SYSTEM SINF_0
  (* Version 1.0, 2023-02-20, eliseu *)
  APPLICATION SINF_0App
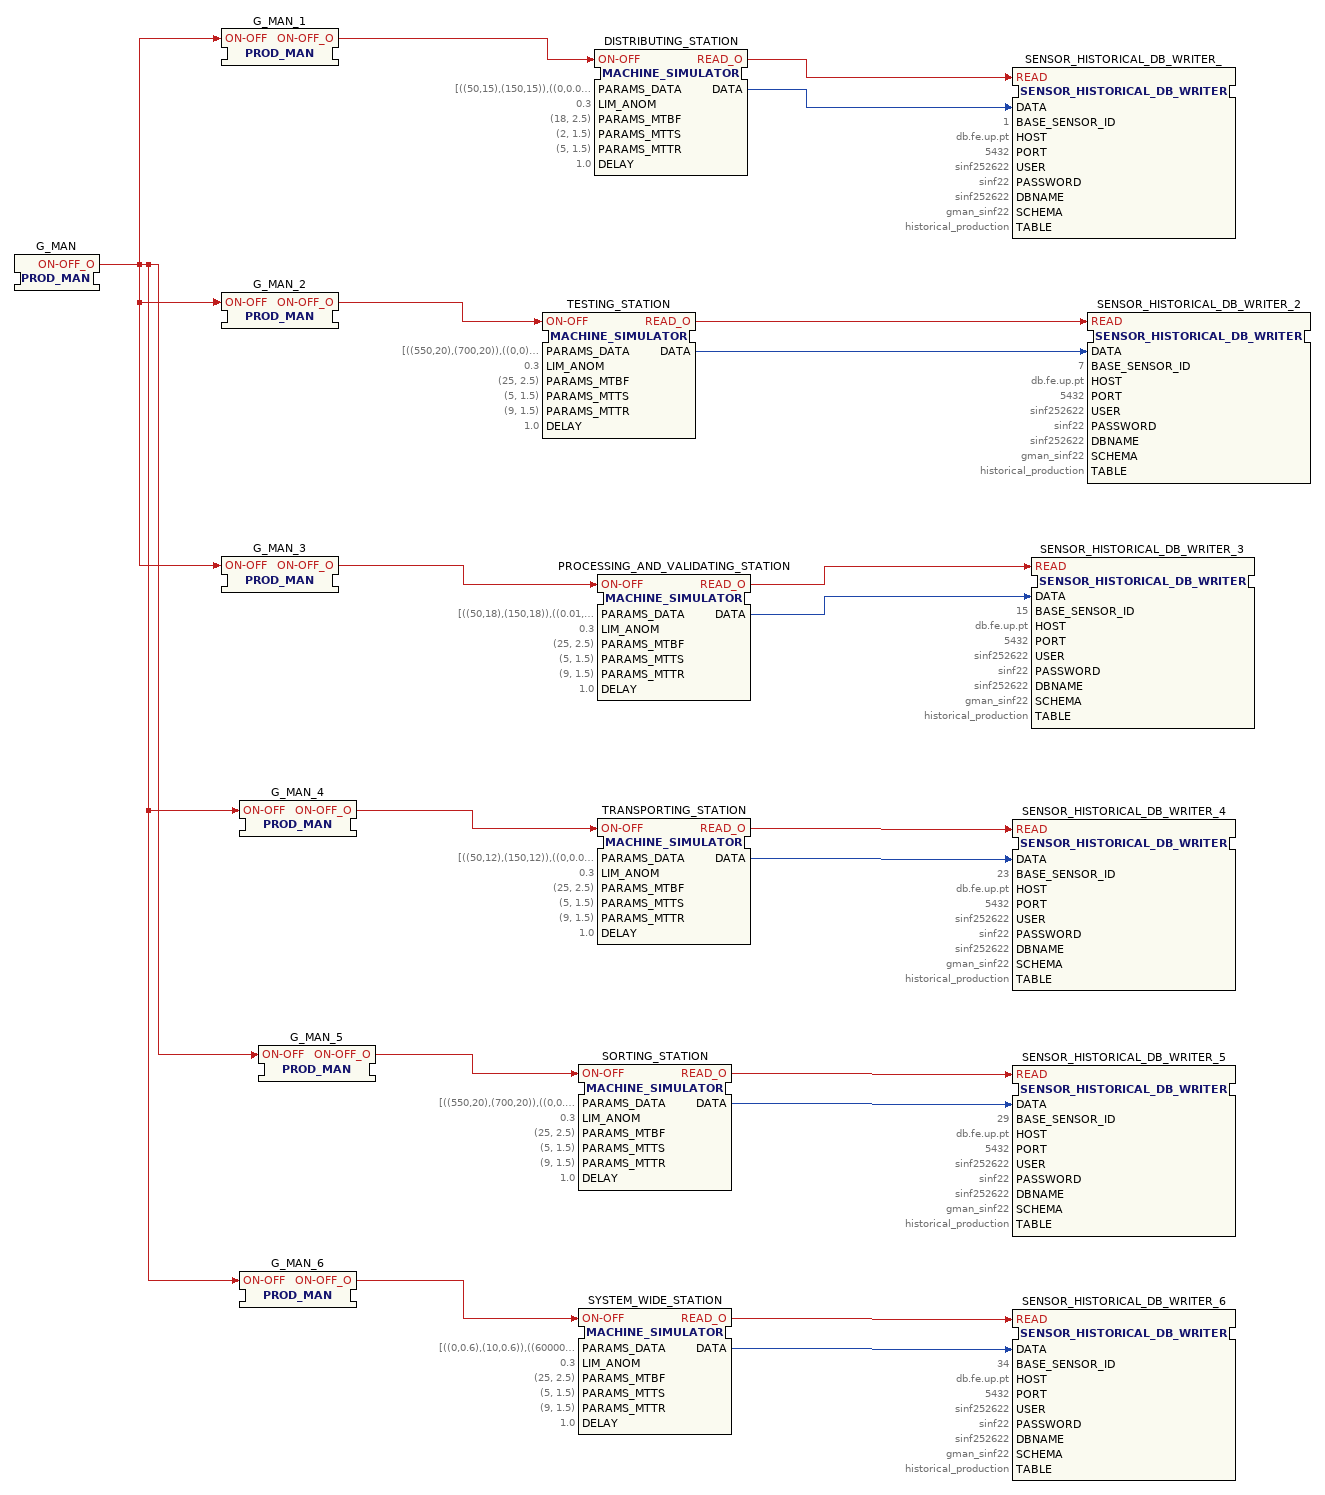
    FBS
      G_MAN_1 : PROD_MAN;
      DISTRIBUTING_STATION : MACHINE_SIMULATOR(PARAMS_DATA := [((50,15),(150,15)),((0,0.05),(3,0.05)),((600000,30000),(800000,30000)),((0.01,0.008),(0.05,0.008)),((2,0.4),(5,0.4)),((293,2.5),(303,2.5))], LIM_ANOM := 0.3, PARAMS_MTBF := (18, 2.5), PARAMS_MTTS := (2, 1.5), PARAMS_MTTR := (5, 1.5), DELAY := 1.0);
      TESTING_STATION : MACHINE_SIMULATOR(PARAMS_DATA := [((550,20),(700,20)),((0,0),(1,0)),((0.2,0.12),(0.8,0.12)),((0,0.05),(3,0.05)),((300,120),(1000,120)),((40,5),(60,5)),((293,2.5),(303,2.5)),((0,0.3),(2,0.3))], LIM_ANOM := 0.3, PARAMS_MTBF := (25, 2.5), PARAMS_MTTS := (5, 1.5), PARAMS_MTTR := (9, 1.5), DELAY := 1.0);
      PROCESSING_AND_VALIDATING_STATION : MACHINE_SIMULATOR(PARAMS_DATA := [((50,18),(150,18)),((0.01,0.012),(0.1,0.012)),((0,0),(1,0)),((0,0.05),(3,0.05)),((2,0.4),(5,0.4)),((333,6),(353,6)),((0.01,0.007),(0.05,0.007)),((500,100),(1000,100))], LIM_ANOM := 0.3, PARAMS_MTBF := (25, 2.5), PARAMS_MTTS := (5, 1.5), PARAMS_MTTR := (9, 1.5), DELAY := 1.0);
      TRANSPORTING_STATION : MACHINE_SIMULATOR(PARAMS_DATA := [((50,12),(150,12)),((0,0.05),(3,0.05)),((2,0.4),(5,0.4)),((333,5),(333,5)),((600000,25000),(800000,25000)),((0.01,0.006),(0.05,0.006))], LIM_ANOM := 0.3, PARAMS_MTBF := (25, 2.5), PARAMS_MTTS := (5, 1.5), PARAMS_MTTR := (9, 1.5), DELAY := 1.0);
      SORTING_STATION : MACHINE_SIMULATOR(PARAMS_DATA := [((550,20),(700,20)),((0,0.05),(3,0.05)),((300,150),(1000,150)),((2,0.35),(5,0.35)),((293,2.5),(303,2.5))], LIM_ANOM := 0.3, PARAMS_MTBF := (25, 2.5), PARAMS_MTTS := (5, 1.5), PARAMS_MTTR := (9, 1.5), DELAY := 1.0);
      SYSTEM_WIDE_STATION : MACHINE_SIMULATOR(PARAMS_DATA := [((0,0.6),(10,0.6)),((600000,30000),(800000,30000)),((40,5),(60,5)),((293,2.5),(303,2.5))], LIM_ANOM := 0.3, PARAMS_MTBF := (25, 2.5), PARAMS_MTTS := (5, 1.5), PARAMS_MTTR := (9, 1.5), DELAY := 1.0);
      G_MAN_2 : PROD_MAN;
      G_MAN_3 : PROD_MAN;
      G_MAN_4 : PROD_MAN;
      G_MAN_5 : PROD_MAN;
      G_MAN_6 : PROD_MAN;
      G_MAN : PROD_MAN;
      SENSOR_HISTORICAL_DB_WRITER_ : SENSOR_HISTORICAL_DB_WRITER(BASE_SENSOR_ID := 1, HOST := db.fe.up.pt, PORT := 5432, USER := sinf252622, PASSWORD := sinf22, DBNAME := sinf252622, SCHEMA := gman_sinf22, TABLE := historical_production);
      SENSOR_HISTORICAL_DB_WRITER_2 : SENSOR_HISTORICAL_DB_WRITER(BASE_SENSOR_ID := 7, HOST := db.fe.up.pt, PORT := 5432, USER := sinf252622, PASSWORD := sinf22, DBNAME := sinf252622, SCHEMA := gman_sinf22, TABLE := historical_production);
      SENSOR_HISTORICAL_DB_WRITER_3 : SENSOR_HISTORICAL_DB_WRITER(BASE_SENSOR_ID := 15, HOST := db.fe.up.pt, PORT := 5432, USER := sinf252622, PASSWORD := sinf22, DBNAME := sinf252622, SCHEMA := gman_sinf22, TABLE := historical_production);
      SENSOR_HISTORICAL_DB_WRITER_4 : SENSOR_HISTORICAL_DB_WRITER(BASE_SENSOR_ID := 23, HOST := db.fe.up.pt, PORT := 5432, USER := sinf252622, PASSWORD := sinf22, DBNAME := sinf252622, SCHEMA := gman_sinf22, TABLE := historical_production);
      SENSOR_HISTORICAL_DB_WRITER_5 : SENSOR_HISTORICAL_DB_WRITER(BASE_SENSOR_ID := 29, HOST := db.fe.up.pt, PORT := 5432, USER := sinf252622, PASSWORD := sinf22, DBNAME := sinf252622, SCHEMA := gman_sinf22, TABLE := historical_production);
      SENSOR_HISTORICAL_DB_WRITER_6 : SENSOR_HISTORICAL_DB_WRITER(BASE_SENSOR_ID := 34, HOST := db.fe.up.pt, PORT := 5432, USER := sinf252622, PASSWORD := sinf22, DBNAME := sinf252622, SCHEMA := gman_sinf22, TABLE := historical_production);
    END_FBS
    EVENT_CONNECTIONS
      G_MAN_1.ON-OFF_O TO DISTRIBUTING_STATION.ON-OFF;
      G_MAN_2.ON-OFF_O TO TESTING_STATION.ON-OFF;
      G_MAN_3.ON-OFF_O TO PROCESSING_AND_VALIDATING_STATION.ON-OFF;
      G_MAN_4.ON-OFF_O TO TRANSPORTING_STATION.ON-OFF;
      G_MAN_5.ON-OFF_O TO SORTING_STATION.ON-OFF;
      G_MAN_6.ON-OFF_O TO SYSTEM_WIDE_STATION.ON-OFF;
      G_MAN.ON-OFF_O TO G_MAN_1.ON-OFF;
      G_MAN.ON-OFF_O TO G_MAN_2.ON-OFF;
      G_MAN.ON-OFF_O TO G_MAN_3.ON-OFF;
      G_MAN.ON-OFF_O TO G_MAN_4.ON-OFF;
      G_MAN.ON-OFF_O TO G_MAN_5.ON-OFF;
      G_MAN.ON-OFF_O TO G_MAN_6.ON-OFF;
      DISTRIBUTING_STATION.READ_O TO SENSOR_HISTORICAL_DB_WRITER_.READ;
      TESTING_STATION.READ_O TO SENSOR_HISTORICAL_DB_WRITER_2.READ;
      SORTING_STATION.READ_O TO SENSOR_HISTORICAL_DB_WRITER_5.READ;
      TRANSPORTING_STATION.READ_O TO SENSOR_HISTORICAL_DB_WRITER_4.READ;
      PROCESSING_AND_VALIDATING_STATION.READ_O TO SENSOR_HISTORICAL_DB_WRITER_3.READ;
      SYSTEM_WIDE_STATION.READ_O TO SENSOR_HISTORICAL_DB_WRITER_6.READ;
    END_CONNECTIONS
    DATA_CONNECTIONS
      DISTRIBUTING_STATION.DATA TO SENSOR_HISTORICAL_DB_WRITER_.DATA;
      TESTING_STATION.DATA TO SENSOR_HISTORICAL_DB_WRITER_2.DATA;
      SORTING_STATION.DATA TO SENSOR_HISTORICAL_DB_WRITER_5.DATA;
      PROCESSING_AND_VALIDATING_STATION.DATA TO SENSOR_HISTORICAL_DB_WRITER_3.DATA;
      SYSTEM_WIDE_STATION.DATA TO SENSOR_HISTORICAL_DB_WRITER_6.DATA;
      TRANSPORTING_STATION.DATA TO SENSOR_HISTORICAL_DB_WRITER_4.DATA;
    END_CONNECTIONS
  END_APPLICATION
  DEVICE FORTE_PC : FORTE_PC(MGR_ID := "localhost:61499")
    {SET_ATTRIBUTE(Profile, HOLOBLOC)} (* device profile *)
    RESOURCE DIN1 : EMB_RES
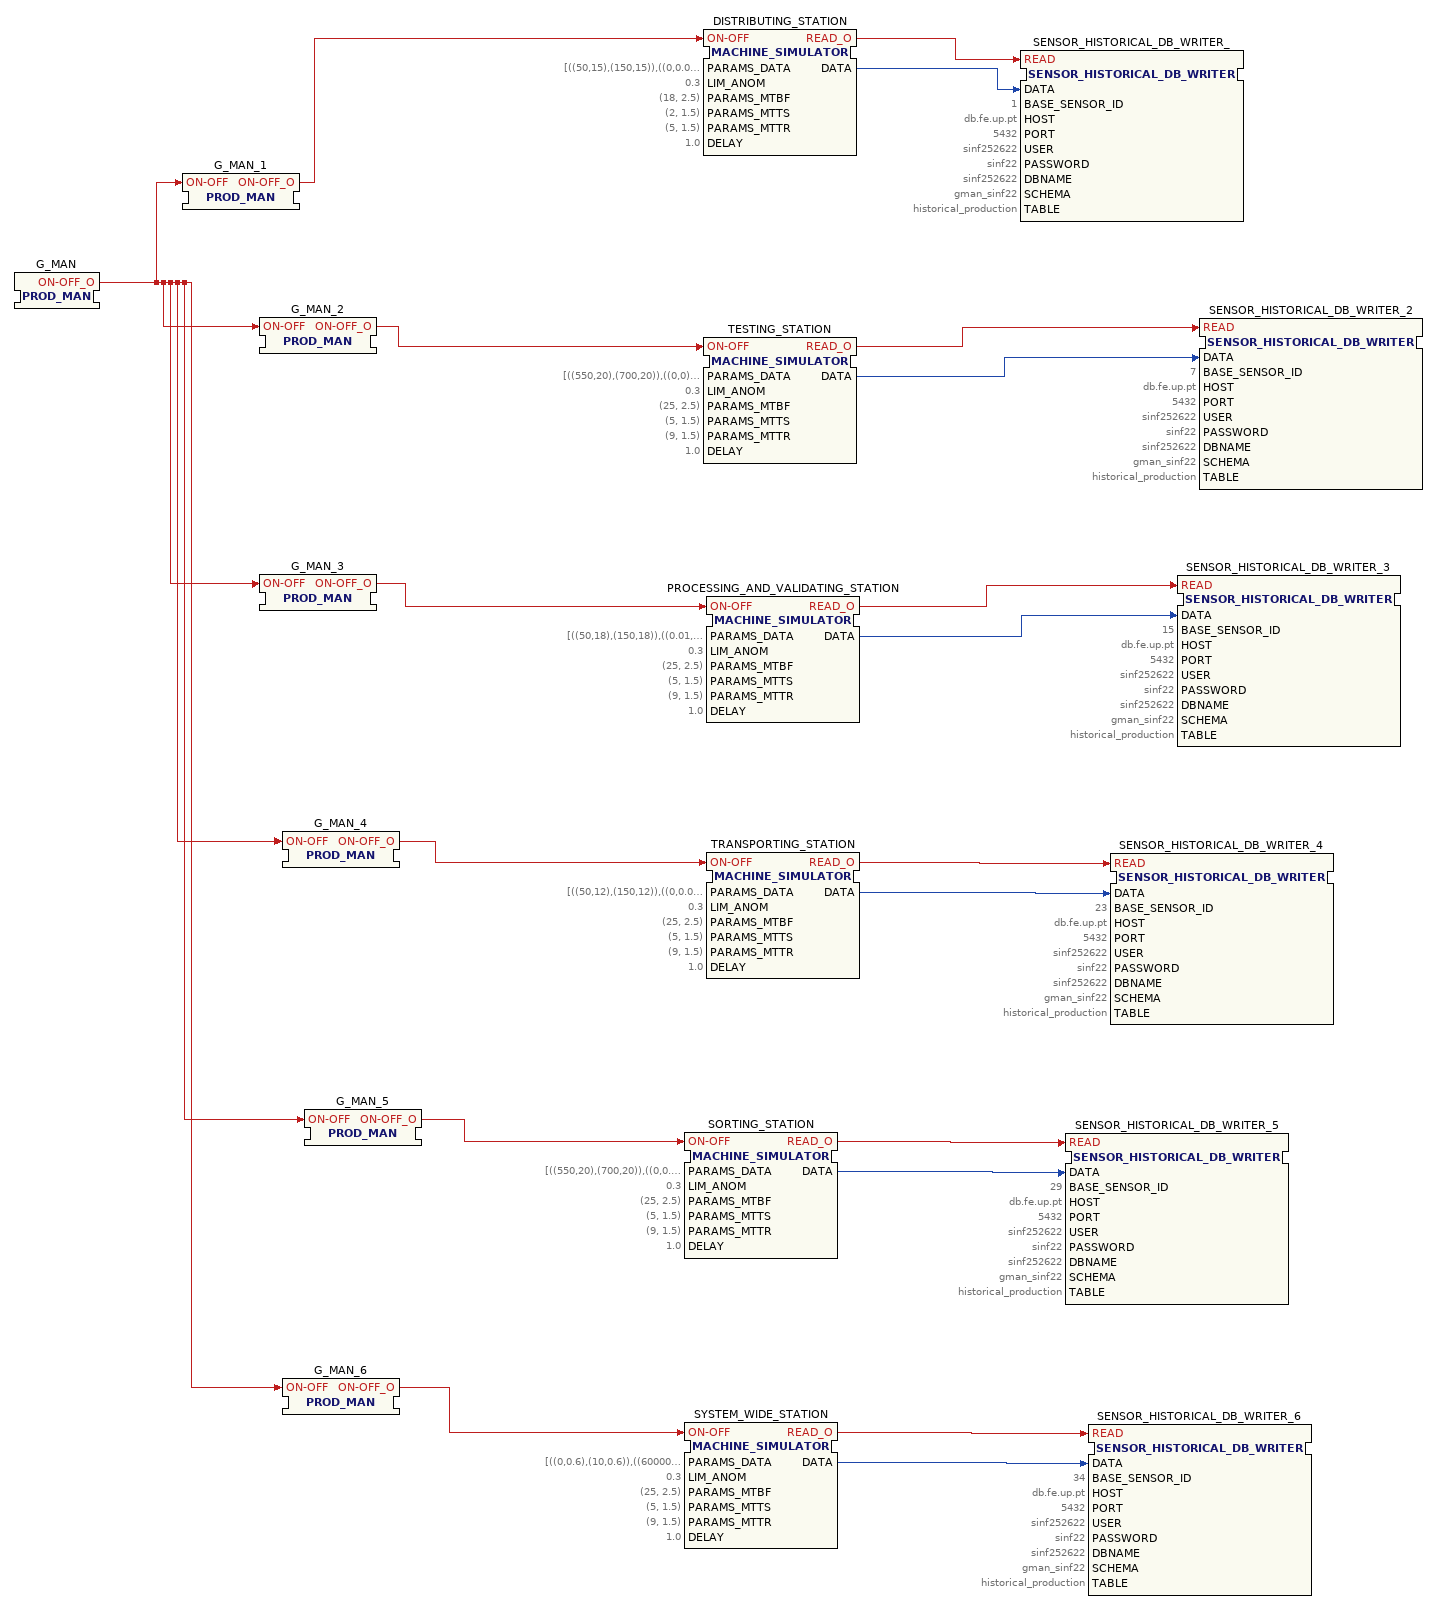
      FBS
        G_MAN_1 : PROD_MAN;
        DISTRIBUTING_STATION : MACHINE_SIMULATOR(PARAMS_DATA := [((50,15),(150,15)),((0,0.05),(3,0.05)),((600000,30000),(800000,30000)),((0.01,0.008),(0.05,0.008)),((2,0.4),(5,0.4)),((293,2.5),(303,2.5))], LIM_ANOM := 0.3, PARAMS_MTBF := (18, 2.5), PARAMS_MTTS := (2, 1.5), PARAMS_MTTR := (5, 1.5), DELAY := 1.0);
        TESTING_STATION : MACHINE_SIMULATOR(PARAMS_DATA := [((550,20),(700,20)),((0,0),(1,0)),((0.2,0.12),(0.8,0.12)),((0,0.05),(3,0.05)),((300,120),(1000,120)),((40,5),(60,5)),((293,2.5),(303,2.5)),((0,0.3),(2,0.3))], LIM_ANOM := 0.3, PARAMS_MTBF := (25, 2.5), PARAMS_MTTS := (5, 1.5), PARAMS_MTTR := (9, 1.5), DELAY := 1.0);
        PROCESSING_AND_VALIDATING_STATION : MACHINE_SIMULATOR(PARAMS_DATA := [((50,18),(150,18)),((0.01,0.012),(0.1,0.012)),((0,0),(1,0)),((0,0.05),(3,0.05)),((2,0.4),(5,0.4)),((333,6),(353,6)),((0.01,0.007),(0.05,0.007)),((500,100),(1000,100))], LIM_ANOM := 0.3, PARAMS_MTBF := (25, 2.5), PARAMS_MTTS := (5, 1.5), PARAMS_MTTR := (9, 1.5), DELAY := 1.0);
        TRANSPORTING_STATION : MACHINE_SIMULATOR(PARAMS_DATA := [((50,12),(150,12)),((0,0.05),(3,0.05)),((2,0.4),(5,0.4)),((333,5),(333,5)),((600000,25000),(800000,25000)),((0.01,0.006),(0.05,0.006))], LIM_ANOM := 0.3, PARAMS_MTBF := (25, 2.5), PARAMS_MTTS := (5, 1.5), PARAMS_MTTR := (9, 1.5), DELAY := 1.0);
        SORTING_STATION : MACHINE_SIMULATOR(PARAMS_DATA := [((550,20),(700,20)),((0,0.05),(3,0.05)),((300,150),(1000,150)),((2,0.35),(5,0.35)),((293,2.5),(303,2.5))], LIM_ANOM := 0.3, PARAMS_MTBF := (25, 2.5), PARAMS_MTTS := (5, 1.5), PARAMS_MTTR := (9, 1.5), DELAY := 1.0);
        SYSTEM_WIDE_STATION : MACHINE_SIMULATOR(PARAMS_DATA := [((0,0.6),(10,0.6)),((600000,30000),(800000,30000)),((40,5),(60,5)),((293,2.5),(303,2.5))], LIM_ANOM := 0.3, PARAMS_MTBF := (25, 2.5), PARAMS_MTTS := (5, 1.5), PARAMS_MTTR := (9, 1.5), DELAY := 1.0);
        G_MAN_2 : PROD_MAN;
        G_MAN_3 : PROD_MAN;
        G_MAN_4 : PROD_MAN;
        G_MAN_5 : PROD_MAN;
        G_MAN_6 : PROD_MAN;
        G_MAN : PROD_MAN;
        SENSOR_HISTORICAL_DB_WRITER_ : SENSOR_HISTORICAL_DB_WRITER(BASE_SENSOR_ID := 1, HOST := db.fe.up.pt, PORT := 5432, USER := sinf252622, PASSWORD := sinf22, DBNAME := sinf252622, SCHEMA := gman_sinf22, TABLE := historical_production);
        SENSOR_HISTORICAL_DB_WRITER_2 : SENSOR_HISTORICAL_DB_WRITER(BASE_SENSOR_ID := 7, HOST := db.fe.up.pt, PORT := 5432, USER := sinf252622, PASSWORD := sinf22, DBNAME := sinf252622, SCHEMA := gman_sinf22, TABLE := historical_production);
        SENSOR_HISTORICAL_DB_WRITER_3 : SENSOR_HISTORICAL_DB_WRITER(BASE_SENSOR_ID := 15, HOST := db.fe.up.pt, PORT := 5432, USER := sinf252622, PASSWORD := sinf22, DBNAME := sinf252622, SCHEMA := gman_sinf22, TABLE := historical_production);
        SENSOR_HISTORICAL_DB_WRITER_4 : SENSOR_HISTORICAL_DB_WRITER(BASE_SENSOR_ID := 23, HOST := db.fe.up.pt, PORT := 5432, USER := sinf252622, PASSWORD := sinf22, DBNAME := sinf252622, SCHEMA := gman_sinf22, TABLE := historical_production);
        SENSOR_HISTORICAL_DB_WRITER_5 : SENSOR_HISTORICAL_DB_WRITER(BASE_SENSOR_ID := 29, HOST := db.fe.up.pt, PORT := 5432, USER := sinf252622, PASSWORD := sinf22, DBNAME := sinf252622, SCHEMA := gman_sinf22, TABLE := historical_production);
        SENSOR_HISTORICAL_DB_WRITER_6 : SENSOR_HISTORICAL_DB_WRITER(BASE_SENSOR_ID := 34, HOST := db.fe.up.pt, PORT := 5432, USER := sinf252622, PASSWORD := sinf22, DBNAME := sinf252622, SCHEMA := gman_sinf22, TABLE := historical_production);
      END_FBS
      EVENT_CONNECTIONS
        G_MAN_1.ON-OFF_O TO DISTRIBUTING_STATION.ON-OFF;
        G_MAN_2.ON-OFF_O TO TESTING_STATION.ON-OFF;
        G_MAN_3.ON-OFF_O TO PROCESSING_AND_VALIDATING_STATION.ON-OFF;
        G_MAN_4.ON-OFF_O TO TRANSPORTING_STATION.ON-OFF;
        G_MAN_5.ON-OFF_O TO SORTING_STATION.ON-OFF;
        G_MAN_6.ON-OFF_O TO SYSTEM_WIDE_STATION.ON-OFF;
        G_MAN.ON-OFF_O TO G_MAN_1.ON-OFF;
        G_MAN.ON-OFF_O TO G_MAN_2.ON-OFF;
        G_MAN.ON-OFF_O TO G_MAN_3.ON-OFF;
        G_MAN.ON-OFF_O TO G_MAN_4.ON-OFF;
        G_MAN.ON-OFF_O TO G_MAN_5.ON-OFF;
        G_MAN.ON-OFF_O TO G_MAN_6.ON-OFF;
        DISTRIBUTING_STATION.READ_O TO SENSOR_HISTORICAL_DB_WRITER_.READ;
        TESTING_STATION.READ_O TO SENSOR_HISTORICAL_DB_WRITER_2.READ;
        SORTING_STATION.READ_O TO SENSOR_HISTORICAL_DB_WRITER_5.READ;
        TRANSPORTING_STATION.READ_O TO SENSOR_HISTORICAL_DB_WRITER_4.READ;
        PROCESSING_AND_VALIDATING_STATION.READ_O TO SENSOR_HISTORICAL_DB_WRITER_3.READ;
        SYSTEM_WIDE_STATION.READ_O TO SENSOR_HISTORICAL_DB_WRITER_6.READ;
      END_CONNECTIONS
      DATA_CONNECTIONS
        DISTRIBUTING_STATION.DATA TO SENSOR_HISTORICAL_DB_WRITER_.DATA;
        TESTING_STATION.DATA TO SENSOR_HISTORICAL_DB_WRITER_2.DATA;
        SORTING_STATION.DATA TO SENSOR_HISTORICAL_DB_WRITER_5.DATA;
        PROCESSING_AND_VALIDATING_STATION.DATA TO SENSOR_HISTORICAL_DB_WRITER_3.DATA;
        SYSTEM_WIDE_STATION.DATA TO SENSOR_HISTORICAL_DB_WRITER_6.DATA;
        TRANSPORTING_STATION.DATA TO SENSOR_HISTORICAL_DB_WRITER_4.DATA;
      END_CONNECTIONS
    END_RESOURCE
  END_DEVICE
  MAPPINGS
    SINF_0App.G_MAN_1 ON FORTE_PC.DIN1.G_MAN_1;
    SINF_0App.DISTRIBUTING_STATION ON FORTE_PC.DIN1.DISTRIBUTING_STATION;
    SINF_0App.TESTING_STATION ON FORTE_PC.DIN1.TESTING_STATION;
    SINF_0App.PROCESSING_AND_VALIDATING_STATION ON FORTE_PC.DIN1.PROCESSING_AND_VALIDATING_STATION;
    SINF_0App.TRANSPORTING_STATION ON FORTE_PC.DIN1.TRANSPORTING_STATION;
    SINF_0App.SORTING_STATION ON FORTE_PC.DIN1.SORTING_STATION;
    SINF_0App.SYSTEM_WIDE_STATION ON FORTE_PC.DIN1.SYSTEM_WIDE_STATION;
    SINF_0App.G_MAN_2 ON FORTE_PC.DIN1.G_MAN_2;
    SINF_0App.G_MAN_3 ON FORTE_PC.DIN1.G_MAN_3;
    SINF_0App.G_MAN_4 ON FORTE_PC.DIN1.G_MAN_4;
    SINF_0App.G_MAN_5 ON FORTE_PC.DIN1.G_MAN_5;
    SINF_0App.G_MAN_6 ON FORTE_PC.DIN1.G_MAN_6;
    SINF_0App.G_MAN ON FORTE_PC.DIN1.G_MAN;
    SINF_0App.SENSOR_HISTORICAL_DB_WRITER_ ON FORTE_PC.DIN1.SENSOR_HISTORICAL_DB_WRITER_;
    SINF_0App.SENSOR_HISTORICAL_DB_WRITER_2 ON FORTE_PC.DIN1.SENSOR_HISTORICAL_DB_WRITER_2;
    SINF_0App.SENSOR_HISTORICAL_DB_WRITER_3 ON FORTE_PC.DIN1.SENSOR_HISTORICAL_DB_WRITER_3;
    SINF_0App.SENSOR_HISTORICAL_DB_WRITER_4 ON FORTE_PC.DIN1.SENSOR_HISTORICAL_DB_WRITER_4;
    SINF_0App.SENSOR_HISTORICAL_DB_WRITER_5 ON FORTE_PC.DIN1.SENSOR_HISTORICAL_DB_WRITER_5;
    SINF_0App.SENSOR_HISTORICAL_DB_WRITER_6 ON FORTE_PC.DIN1.SENSOR_HISTORICAL_DB_WRITER_6;
  END_MAPPINGS
  SEGMENTS
    Ethernet : Ethernet;
  END_SEGMENTS
  LINKS
    FORTE_PC => Ethernet;
  END_LINKS
END_SYSTEM
